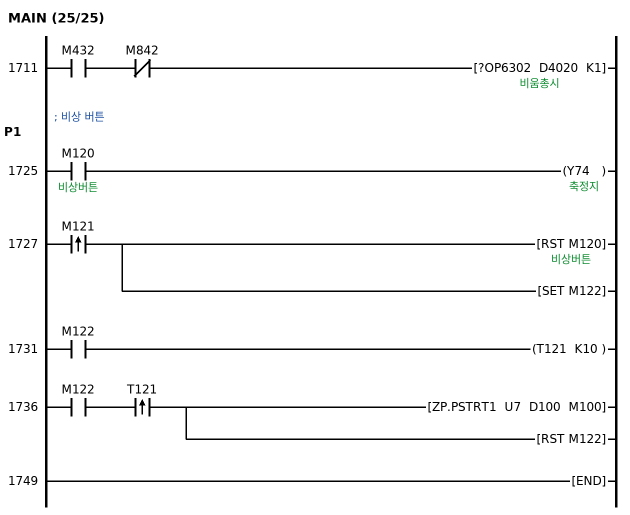
[picture p24: ladder of MAIN, rungs at steps 1711 to 1749]
1711  LD      M432
      ANI     M842
      ?OP6302 D4020 K1
; 비상 버튼
      P1
1725  LD      M120  ; 비상버튼
      OUT     Y74  ; 축정지
1727  LDP     M121
      RST     M120  ; 비상버튼
      SET     M122
1731  LD      M122
      OUT     T121 K10
1736  LD      M122
      ANDP    T121
      ZP.PSTRT1 U7 D100 M100
      RST     M122
1749  END
END_PROGRAM

PROGRAM OUTPUT
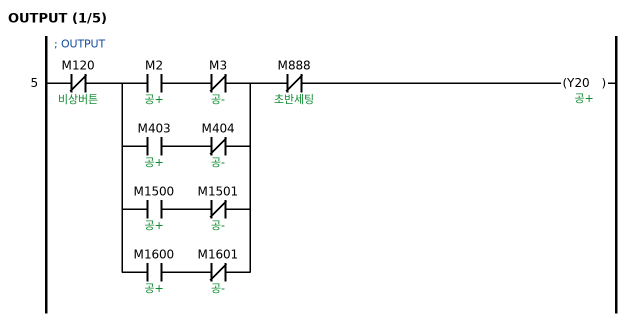
; OUTPUT
5     LDI     M120  ; 비상버튼
      LD      M2  ; 공+
      ANI     M3  ; 공-
      LD      M403  ; 공+
      ANI     M404  ; 공-
      ORB
      LD      M1500  ; 공+
      ANI     M1501  ; 공-
      ORB
      LD      M1600  ; 공+
      ANI     M1601  ; 공-
      ORB
      ANB
      ANI     M888  ; 초반세팅
      OUT     Y20  ; 공+
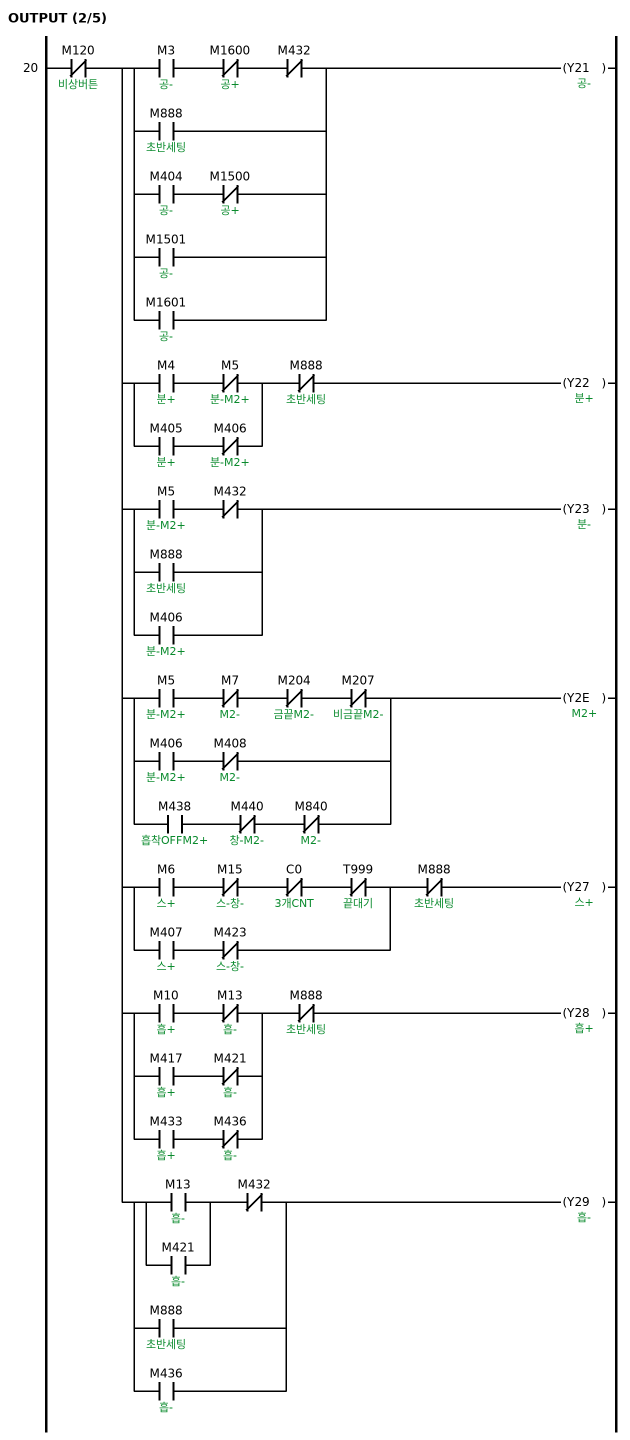
20    LDI     M120  ; 비상버튼
      MPS
      LD      M3  ; 공-
      ANI     M1600  ; 공+
      ANI     M432
      OR      M888  ; 초반세팅
      LD      M404  ; 공-
      ANI     M1500  ; 공+
      ORB
      OR      M1501  ; 공-
      OR      M1601  ; 공-
      ANB
      OUT     Y21  ; 공-
      MRD
      LD      M4  ; 분+
      ANI     M5  ; 분-M2+
      LD      M405  ; 분+
      ANI     M406  ; 분-M2+
      ORB
      ANB
      ANI     M888  ; 초반세팅
      OUT     Y22  ; 분+
      MRD
      LD      M5  ; 분-M2+
      ANI     M432
      OR      M888  ; 초반세팅
      OR      M406  ; 분-M2+
      ANB
      OUT     Y23  ; 분-
      MRD
      LD      M5  ; 분-M2+
      ANI     M7  ; M2-
      ANI     M204  ; 금끝M2-
      ANI     M207  ; 비금끝M2-
      LD      M406  ; 분-M2+
      ANI     M408  ; M2-
      ORB
      LD      M438  ; 흡착OFFM2+
      ANI     M440  ; 창-M2-
      ANI     M840  ; M2-
      ORB
      ANB
      OUT     Y2E  ; M2+
      MRD
      LD      M6  ; 스+
      ANI     M15  ; 스-창-
      ANI     C0  ; 3개CNT
      ANI     T999  ; 끝대기
      LD      M407  ; 스+
      ANI     M423  ; 스-창-
      ORB
      ANB
      ANI     M888  ; 초반세팅
      OUT     Y27  ; 스+
      MRD
      LD      M10  ; 흡+
      ANI     M13  ; 흡-
      LD      M417  ; 흡+
      ANI     M421  ; 흡-
      ORB
      LD      M433  ; 흡+
      ANI     M436  ; 흡-
      ORB
      ANB
      ANI     M888  ; 초반세팅
      OUT     Y28  ; 흡+
      MPP
      LD      M13  ; 흡-
      OR      M421  ; 흡-
      ANI     M432
      OR      M888  ; 초반세팅
      OR      M436  ; 흡-
      ANB
      OUT     Y29  ; 흡-
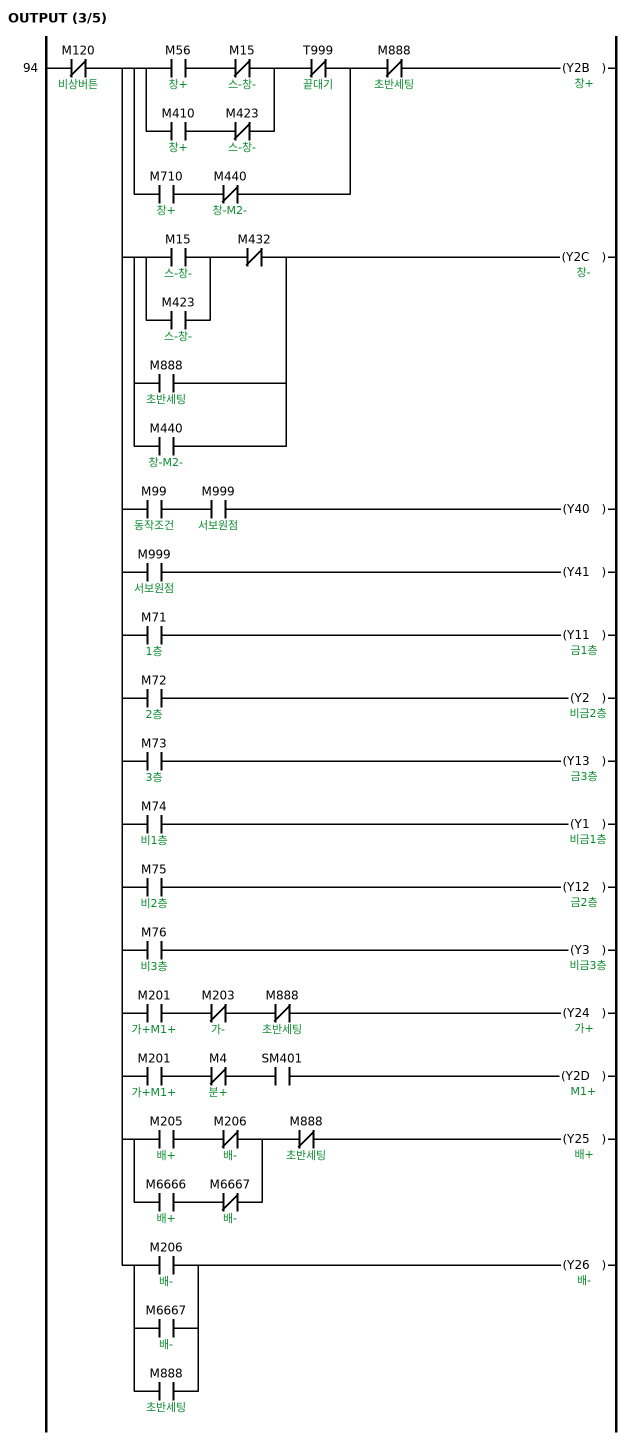
94    LDI     M120  ; 비상버튼
      MPS
      LD      M56  ; 창+
      ANI     M15  ; 스-창-
      LD      M410  ; 창+
      ANI     M423  ; 스-창-
      ORB
      ANI     T999  ; 끝대기
      LD      M710  ; 창+
      ANI     M440  ; 창-M2-
      ORB
      ANB
      ANI     M888  ; 초반세팅
      OUT     Y2B  ; 창+
      MRD
      LD      M15  ; 스-창-
      OR      M423  ; 스-창-
      ANI     M432
      OR      M888  ; 초반세팅
      OR      M440  ; 창-M2-
      ANB
      OUT     Y2C  ; 창-
      MRD
      AND     M99  ; 동작조건
      AND     M999  ; 서보원점
      OUT     Y40
      MRD
      AND     M999  ; 서보원점
      OUT     Y41
      MRD
      AND     M71  ; 1층
      OUT     Y11  ; 금1층
      MRD
      AND     M72  ; 2층
      OUT     Y2  ; 비금2층
      MRD
      AND     M73  ; 3층
      OUT     Y13  ; 금3층
      MRD
      AND     M74  ; 비1층
      OUT     Y1  ; 비금1층
      MRD
      AND     M75  ; 비2층
      OUT     Y12  ; 금2층
      MRD
      AND     M76  ; 비3층
      OUT     Y3  ; 비금3층
      MRD
      AND     M201  ; 가+M1+
      ANI     M203  ; 가-
      ANI     M888  ; 초반세팅
      OUT     Y24  ; 가+
      MRD
      AND     M201  ; 가+M1+
      ANI     M4  ; 분+
      AND     SM401
      OUT     Y2D  ; M1+
      MRD
      LD      M205  ; 배+
      ANI     M206  ; 배-
      LD      M6666  ; 배+
      ANI     M6667  ; 배-
      ORB
      ANB
      ANI     M888  ; 초반세팅
      OUT     Y25  ; 배+
      MPP
      LD      M206  ; 배-
      OR      M6667  ; 배-
      OR      M888  ; 초반세팅
      ANB
      OUT     Y26  ; 배-
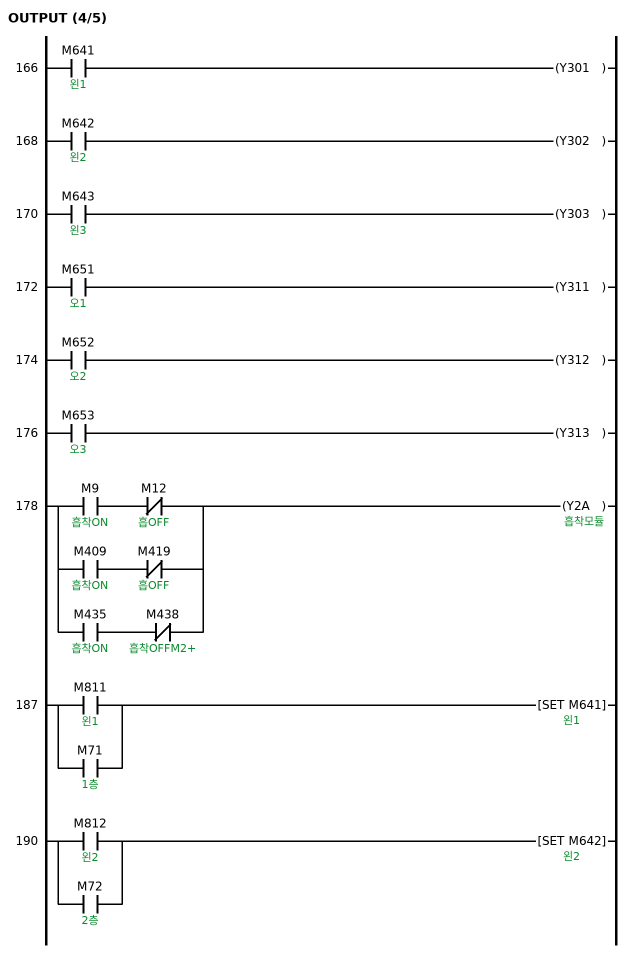
166   LD      M641  ; 왼1
      OUT     Y301
168   LD      M642  ; 왼2
      OUT     Y302
170   LD      M643  ; 왼3
      OUT     Y303
172   LD      M651  ; 오1
      OUT     Y311
174   LD      M652  ; 오2
      OUT     Y312
176   LD      M653  ; 오3
      OUT     Y313
178   LD      M9  ; 흡착ON
      ANI     M12  ; 흡OFF
      LD      M409  ; 흡착ON
      ANI     M419  ; 흡OFF
      ORB
      LD      M435  ; 흡착ON
      ANI     M438  ; 흡착OFFM2+
      ORB
      OUT     Y2A  ; 흡착모듈
187   LD      M811  ; 왼1
      OR      M71  ; 1층
      SET     M641  ; 왼1
190   LD      M812  ; 왼2
      OR      M72  ; 2층
      SET     M642  ; 왼2
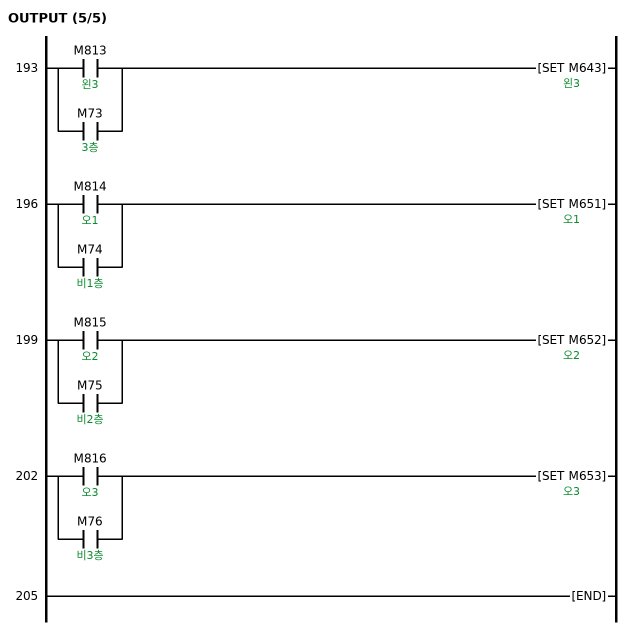
193   LD      M813  ; 왼3
      OR      M73  ; 3층
      SET     M643  ; 왼3
196   LD      M814  ; 오1
      OR      M74  ; 비1층
      SET     M651  ; 오1
199   LD      M815  ; 오2
      OR      M75  ; 비2층
      SET     M652  ; 오2
202   LD      M816  ; 오3
      OR      M76  ; 비3층
      SET     M653  ; 오3
205   END
END_PROGRAM

// device comments not shown above
X5  ; 가+
X0C  ; X7C
X0E  ; 창+
M18  ; 종료
M51  ; 비금1층
M52  ; 비금2층
M53  ; 비금3층
M61  ; 금1층
M62  ; 금2층
M63  ; 금3층
M67  ; 창-
M111  ; 원점복귀
M119  ; 비상 중지
M222  ; 가공반복
M333  ; 시작
M481  ; 왼쪽1층
M556  ; 비금1층
M557  ; 비금2층
M558  ; 비금3층
M667  ; 금속1층
M668  ; 금속2층
M669  ; 금속3층
M1002  ; 고속원점
M1006  ; 수동동작
M1111  ; 원점복귀
M2000  ; 소재흡착
M2002  ; 2층
M2003  ; 3층
M2004  ; 흡착ONOFF
M2005  ; 흡착전진
M2006  ; 흡착후진
M2007  ; 흡착위치
M2008  ; 이송위치
M2055  ; 전진완
M2066  ; 후진완
T200  ; 가공대기
D300  ; 시간총합
